Fanuc KAREL source: kb00078.KL

PROGRAM KB00078
%STACKSIZE=65535
%PRIORITY=65535
%NOLOCKGROUP
VAR
P1 : FILE
RESULT : INTEGER
BEGIN
RESULT=GET_FILE_POS(P1)
END KB00078
